FUNCTION_BLOCK Recipe2 (* Basic Function Block Type *)
  (* Standard: 61499-2 *)
  (* Version 0.0, 10/11/2026, macie, nxtControl GmBH, Template *)
  PACKAGE Main;
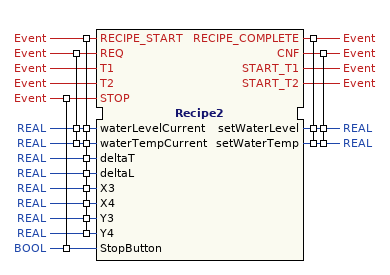
  EVENT_INPUT
    RECIPE_START WITH waterLevelCurrent, waterTempCurrent, deltaT, deltaL, X3, X4, Y3, Y4; (* Initialization Request *)
    REQ WITH waterLevelCurrent, waterTempCurrent; (* Normal Execution Request *)
    T1;
    T2;
    STOP WITH StopButton;
  END_EVENT
  EVENT_OUTPUT
    RECIPE_COMPLETE WITH setWaterLevel, setWaterTemp; (* Initialization Confirm *)
    CNF WITH setWaterLevel, setWaterTemp; (* Execution Confirmation *)
    START_T1;
    START_T2;
  END_EVENT
  VAR_INPUT
    waterLevelCurrent : REAL;
    waterTempCurrent : REAL; (* Input event qualifier *)
    deltaT : REAL;
    deltaL : REAL;
    X3 : REAL;
    X4 : REAL;
    Y3 : REAL;
    Y4 : REAL;
    StopButton : BOOL;
  END_VAR
  VAR_OUTPUT
    setWaterLevel : REAL; (* Output event qualifier *)
    setWaterTemp : REAL;
  END_VAR
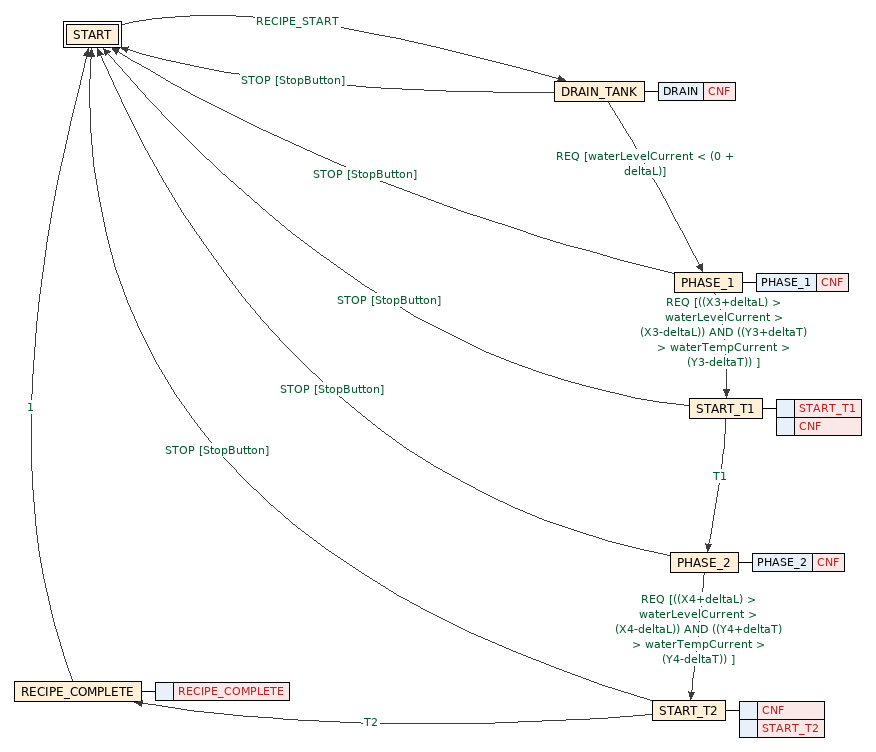
  EC_STATES
    START; (* Initial State *)
    DRAIN_TANK : DRAIN -> CNF;
    PHASE_1 : PHASE_1 -> CNF;
    PHASE_2 : PHASE_2 -> CNF;
    START_T2 : -> CNF, -> START_T2;
    RECIPE_COMPLETE : -> RECIPE_COMPLETE;
    START_T1 : -> START_T1, -> CNF;
  END_STATES
  EC_TRANSITIONS
    START TO DRAIN_TANK := RECIPE_START;
    DRAIN_TANK TO PHASE_1 := REQ [waterLevelCurrent < (0 + deltaL)];
    PHASE_1 TO START_T1 := REQ [((X3+deltaL) > waterLevelCurrent > (X3-deltaL)) AND ((Y3+deltaT) > waterTempCurrent > (Y3-deltaT)) ];
    PHASE_2 TO START_T2 := REQ [((X4+deltaL) > waterLevelCurrent > (X4-deltaL)) AND ((Y4+deltaT) > waterTempCurrent > (Y4-deltaT)) ];
    RECIPE_COMPLETE TO START := 1;
    START_T1 TO PHASE_2 := T1;
    START_T2 TO RECIPE_COMPLETE := T2;
    DRAIN_TANK TO START := STOP [StopButton];
    PHASE_1 TO START := STOP [StopButton];
    START_T1 TO START := STOP [StopButton];
    PHASE_2 TO START := STOP [StopButton];
    START_T2 TO START := STOP [StopButton];
  END_TRANSITIONS
  ALGORITHM INIT IN ST: (* Initialization algorithm *)
;
  END_ALGORITHM
  ALGORITHM REQ IN ST: (* Normally executed algorithm *)
;
  END_ALGORITHM
  ALGORITHM DRAIN IN ST:
;
setWaterLevel := 0;
setWaterTemp := 0;
  END_ALGORITHM
  ALGORITHM PHASE_1 IN ST:
;
setWaterLevel := X3;
setWaterTemp := Y3;
  END_ALGORITHM
  ALGORITHM PHASE_2 IN ST:
;
setWaterLevel := X4;
setWaterTemp := Y4;
  END_ALGORITHM
END_FUNCTION_BLOCK
